(*
SPDX-FileCopyrightText: © 2026 Oleksandr Tiutyk <trofimich@gmail.com>
SPDX-License-Identifier: MIT
License: https://opensource.org/license/mit
*)

(*!
<summary>Defines a condition that combines child conditions with a logical AND or OR operator.</summary>
*)

INTERFACE ICompositeCondition EXTENDS ICondition

(*!
<summary>Appends a child condition to this composite condition.</summary>
<description>
Rejects null references, cycles and conditions already attached to another parent.
The standard implementation also rejects duplicate slots, validates fixed workflow association and requires
the parent chain and owning workflow to be PASSIVE_READY before mutation. Child storage remains borrowed.
</description>
<param name="condition">Child condition to append.</param>
*)
METHOD AddChildCondition
VAR_INPUT
	condition : ICondition;
END_VAR
END_METHOD

(*!
<summary>Gets or sets the logical operator (AND_ or OR_) used to combine child conditions.</summary>
*)
PROPERTY LogicalOperator : LOGICAL_OPERATOR
GET
END_GET
SET
END_SET
END_PROPERTY

END_INTERFACE

(* stored: Version 1.1.0.1
   Itf ICompositeCondition: Id {5071de02-a2b1-4cba-93bf-27c0973efb35}
   Method AddChildCondition: Id {dc921a49-202f-47b9-adb5-2f8dad5d5097}
   Property LogicalOperator: Id {30ffe6f4-aae4-4362-aacc-960e71565572}
   Get Get: Id {e3fc3c86-048d-4ff0-a309-84663d1eab60}
   Set Set: Id {f9275521-91e9-460d-b8b6-72fa668ebc4c} *)
